(* IEC 61131-3 sources: llm-plc-st-eval/data/definitivo/gpt-4o-2024-08-06/C8/zero_shot, 3 files *)

(* ---- ejec_1.st ---- *)
```pascal
FUNCTION_BLOCK FB_Valvula
VAR
    nivelAlto : BOOL; // Entrada: indica si el nivel es alto
    valvula : BOOL;   // Salida: controla la válvula
    T1 : TON;         // Temporizador TON
END_VAR

// Inicialización del temporizador
T1(IN := nivelAlto, PT := T#5S);

// Control de la válvula basado en el temporizador
valvula := T1.Q;
END_FUNCTION_BLOCK
```

Este código en Structured Text (ST) implementa el comportamiento descrito en el Ladder Diagram, utilizando un temporizador TON y controlando la salida `valvula` según el estado del temporizador.

(* ---- ejec_2.st ---- *)
```pascal
FUNCTION_BLOCK FB_Valvula
VAR
    nivelAlto : BOOL; // Entrada: indica si el nivel es alto
    valvula : BOOL;   // Salida: controla la válvula
    T1 : TON;         // Temporizador TON
END_VAR

// Asignación del tiempo preestablecido del temporizador
T1(IN := nivelAlto, PT := T#5S);

// La salida de la válvula se activa si el temporizador ha alcanzado el tiempo preestablecido
valvula := T1.Q;
END_FUNCTION_BLOCK
```

(* ---- ejec_3.st ---- *)
```pascal
FUNCTION_BLOCK FB_Valvula
VAR
    nivelAlto : BOOL; // Entrada: indica si el nivel es alto
    valvula : BOOL;   // Salida: controla la válvula
    T1 : TON;         // Temporizador TON
END_VAR

// Inicialización del temporizador
T1(IN := nivelAlto, PT := T#5S);

// Asignación de la salida de la válvula
valvula := T1.Q;
```

Este código en Structured Text (ST) implementa el comportamiento descrito en el Ladder Diagram, utilizando un temporizador TON para controlar la salida `valvula` basada en la entrada `nivelAlto`.
